{attribute 'Tc2GvlVarNames'}
VAR_GLOBAL

END_VAR

(* stored: Version 1.1.0.1, ProductVersion 3.1.4024.15
   GVL GVL_Gr02Init: Id {a393a1f9-2a41-450b-9671-e0508acb5295} *)
